(*
SPDX-FileCopyrightText: c 2026 Oleksandr Tiutyk <trofimich@gmail.com>
SPDX-License-Identifier: MIT
License: https://opensource.org/license/mit
*)

(*!
<summary>Checks random scaling and a single-point interval.</summary>
<description>
Owns a generator used by one PLC task. Each run checks the same bounds against fresh samples.
The runner binds assertions to the instance address. Keep the instance at that address for its run.
</description>
*)

{attribute 'no_assign'}
{attribute 'no_explicit_call' := 'do not call this function block directly'}
FUNCTION_BLOCK RandomRangeTest EXTENDS TOF_Testing.SingleCycleTest
VAR_STAT
	{attribute 'hide'}
	_ClassName : STRING := __POUNAME();
END_VAR
VAR
	_Random : TOF_Core.Random;
END_VAR

//! <summary>Checks a single-point range and samples an inclusive interval.</summary>
METHOD PROTECTED ExecuteTest
VAR
	value : LREAL;
	i : INT;
END_VAR
value := _Random.GetInRange(minValue := LREAL#-7.5, maxValue := LREAL#-7.5);
Assert.ThatLongReal(
	actual := value,
	message := "A single-point range must return its bound"
).ToBe(expected := LREAL#-7.5);

FOR i := 1 TO 21 DO
	value := _Random.GetInRange(minValue := LREAL#100.0, maxValue := LREAL#200.0);
	Assert.ThatLongReal(
		actual := value,
		message := "GetInRange sample below 100"
	).IsGreaterThanOrEquals(expected := LREAL#100.0);
	Assert.ThatLongReal(
		actual := value,
		message := "GetInRange sample above 200"
	).IsLessThanOrEquals(expected := LREAL#200.0);
END_FOR
END_METHOD

//! <summary>Borrows the concrete class name. Callers must not modify it.</summary>
{attribute 'monitoring' := 'call'}
PROPERTY ClassName : REFERENCE TO STRING
GET
ClassName REF= _ClassName;
END_GET
END_PROPERTY

//! <summary>Borrows the compiler-initialized namespace name. Callers must not modify it.</summary>
{attribute 'monitoring' := 'call'}
PROPERTY NamespaceName : REFERENCE TO STRING
GET
NamespaceName REF= CurrentNamespace.Name;
END_GET
END_PROPERTY

//! <summary>Reports the concrete instance size in bytes.</summary>
{attribute 'monitoring' := 'call'}
PROPERTY SelfSize : ULINT
GET
SelfSize := XSIZEOF(THIS^);
END_GET
END_PROPERTY

END_FUNCTION_BLOCK

(* stored: Version 1.1.0.1
   POU RandomRangeTest: Id {5add9fe6-8949-468d-810d-3c825c4cb768}, SpecialFunc None
   Method ExecuteTest: Id {725e6b80-50b1-41aa-9d4f-11fdc2e3ad75}
   Property ClassName: Id {9255680a-e814-437d-b18b-d3511be2031c}
   Get Get: Id {b33b3207-5386-4868-beb5-998b28eaa25d}
   Property NamespaceName: Id {1f80554d-ac78-4dd6-bccf-241e8d56379b}
   Get Get: Id {f9593dfa-3baf-4782-928c-b687fa58c71a}
   Property SelfSize: Id {8dfbe9e1-337c-4bdc-89ba-d245d894582d}
   Get Get: Id {bdb5698d-fb64-4d21-bc66-4eff730b312d} *)
